(* IEC 61131-3 sources: rusty/compiler/plc_cfc/fixtures/blocks/reference, 3 files *)

(* ---- addInto.st ---- *)
FUNCTION addInto : DINT
    VAR_INPUT
        delta : DINT;
    END_VAR
    VAR_IN_OUT
        acc : DINT;
    END_VAR
    acc := acc + delta;
    addInto := acc;
END_FUNCTION

(* ---- doNothing.st ---- *)
FUNCTION doNothing
VAR_INPUT
    in: DINT;
END_VAR
VAR_OUTPUT
    out: DINT;
END_VAR

// does nothing, alternatively does something but returns no value other than the VAR_OUTPUT variable
END_FUNCTION

FUNCTION doNothing2 : INT
VAR_INPUT
    in: DINT;
END_VAR

END_FUNCTION

(* ---- myAdd.st ---- *)
FUNCTION myAdd : INT
    VAR_INPUT
        in1, in2: DINT;
    END_VAR

    VAR_OUTPUT
        myAddDoubled: DINT;
    END_VAR

    myAdd := in1 + in2;
    myAddDoubled := (in1 + in2) * 2;
END_FUNCTION
